// TIA Portal project "Project5" (V19)

(* hardware
DEVICE "S7-1500/ET200MP station_1"  S7-1500 station
   slot 0: "Rail_0"  Rack  6ES7 590-1***0-0AA0
   slot 1: "PLC_1"  CPU 1511C-1 PN  6ES7 511-1CK01-0AB0  V2.9
      slot 3: "CPU display_1"  6ES7591-1AA00-0AA0
      slot 32768: "PROFINET interface_1"  X1
         slot 32769: "Port_1"  X1 P1
         slot 32770: "Port_2"  X1 P2
      slot 34817: "Virtual CP interface port_1"  Virtual CP interface port  Virtual CP interface port
*)

// ===== PLC "PLC_1"  CPU 1511C-1 PN =====

VAR_GLOBAL   // PLC tag table "Default tag table"
   "Tag_1" AT %MW10 : Word;
   "Tag_2" AT %MD10 : DInt;
   "Tag_3" AT %MD20 : Real;
   "System_Byte" AT %MB100 : Byte;
   "FirstScan" AT %M100.0 : Bool;
   "DiagStatusUpdate" AT %M100.1 : Bool;
   "AlwaysTRUE" AT %M100.2 : Bool;
   "AlwaysFALSE" AT %M100.3 : Bool;
   "System_Byte(1)" AT %MB1 : Byte;
   "Clock_Byte" AT %MB100 : Byte;
   "Clock_10Hz" AT %M100.0 : Bool;
   "Clock_5Hz" AT %M100.1 : Bool;
   "Clock_2.5Hz" AT %M100.2 : Bool;
   "Clock_2Hz" AT %M100.3 : Bool;
   "Clock_1.25Hz" AT %M100.4 : Bool;
   "Clock_1Hz" AT %M100.5 : Bool;
   "Clock_0.625Hz" AT %M100.6 : Bool;
   "Clock_0.5Hz" AT %M100.7 : Bool;
   "Tag_4" AT %MW200 : Word;
   "Tag_5" AT %MW202 : Word;
   "Tag_6" AT %MD202 : Real;
END_VAR

DATA_BLOCK "FB_Motor_Speed_Calc_DB"   // DB1
{ S7_Optimized_Access := 'TRUE' }
VERSION : 0.1
// stored: InstanceOfName FB_Motor_Speed_Calc
"FB_Motor_Speed_Calc"
BEGIN
END_DATA_BLOCK

DATA_BLOCK "FB_Motor_Speed_Calc_Max_DB"   // DB3
{ S7_Optimized_Access := 'TRUE' }
VERSION : 0.2
// stored: InstanceOfName FB_Motor_Speed_Calc_Max
"FB_Motor_Speed_Calc_Max"
BEGIN
END_DATA_BLOCK

FUNCTION_BLOCK "FB_Motor_Speed_Calc"   // FB1, SCL
{ S7_Optimized_Access := 'TRUE' }
VERSION : 0.1
   VAR_INPUT
      Current_HSC_Count : DInt;   // Current value of the high-speed counter (e.g., LADDR#272)
      Run_Calculation : Bool;   // Trigger to run the calculation (e.g., driven by a 1s clock or OB35)
      Measurement_Interval_ms : Real := 1000.0;   // The fixed time interval for measurement (e.g., 1000.0 ms = 1 second)
      Pulses_Per_Revolution : Real := 1.0;   // Number of pulses generated by the sensor per one revolution (User specified 1)
   END_VAR
   VAR_OUTPUT
      RPM_Out : Real;   // Calculated motor speed in Revolutions Per Minute
   END_VAR
   VAR
      Previous_Count : DInt;   // Internal memory to store the count from the last calculation cycle (STATIC)
   END_VAR
   VAR_TEMP
      Time_Interval_s : Real;
      Delta_Count : Real;
   END_VAR
BEGIN
       // ----------------------------------------------------------------------
       // Speed Calculation Logic (Delta Count Method)
       // Runs only when the 'Run_Calculation' trigger is true (e.g., once every second)
       // Formula: RPM = (Delta_Count / Time_Interval_s) * (60.0 / PPR)
       // ----------------------------------------------------------------------

       IF #Run_Calculation THEN

           // 1. Calculate the change in count (Delta_Count)
           // DINT is used for counters. We convert to REAL for calculation accuracy.
           // We must handle the case where the counter may reset (Current < Previous),
           // although for modern PLCs reading a DINT HSC value, this is less likely 
           // to happen within a short interval.

           // Calculate the difference between the current count and the count from the last cycle

           // Check for potential counter rollover (Current_HSC_Count < Previous_Count)
           // If it rolls over, the difference will be negative, and the magnitude will be large,
           // but typically the HSC configuration handles this by resetting to 0. 
           // Assuming a standard incremental count:
           #Delta_Count := DINT_TO_REAL(#Current_HSC_Count -#Previous_Count);

           // 2. Convert the measurement interval from milliseconds to seconds
           #Time_Interval_s := #Measurement_Interval_ms / 1000.0;

           // 3. Check for division by zero (should not happen if Measurement_Interval_ms > 0)
           IF #Time_Interval_s > 0.0 AND #Pulses_Per_Revolution > 0.0 THEN

               // Calculate the speed in RPM
               // (Counts/second) * 60 = Counts/minute
               // (Counts/minute) / PPR = Revolutions/minute (RPM)
               #RPM_Out := (#Delta_Count / #Time_Interval_s) * (60.0 /#Pulses_Per_Revolution);

           ELSE
               #RPM_Out := 0.0;
           END_IF;

           // 4. Store the current count for the next calculation cycle
           #Previous_Count :=#Current_HSC_Count;

       END_IF;
END_FUNCTION_BLOCK

FUNCTION_BLOCK "FB_Motor_Speed_Calc_Max"   // FB2, SCL
{ S7_Optimized_Access := 'TRUE' }
VERSION : 0.2
   VAR_INPUT
      Current_HSC_Count : DInt;   // Current value of the high-speed counter
      Run_Calculation : Bool;   // Trigger to run the calculation (e.g., driven by a 1s clock or OB35)
      Reset_Max_RPM : Bool;   // New input: Use a momentary pulse to reset Max_RPM_Out to 0.0
      Measurement_Interval_ms : Real := 1000.0;   // The fixed time interval for measurement (e.g., 1000.0 ms = 1 second)
      Pulses_Per_Revolution : Real := 1.0;   // Number of pulses generated by the sensor per one revolution
   END_VAR
   VAR_OUTPUT
      RPM_Out : Real;   // Calculated current motor speed in Revolutions Per Minute
      Max_RPM_Out : Real;   // Output: Stores the highest RPM achieved since the last reset
   END_VAR
   VAR
      Previous_Count : DInt;   // Internal memory to store the count from the last calculation cycle (STATIC)
      s_Max_RPM_Value : Real;   // STATIC: Internal memory to persistently store the maximum RPM achieved. Initialized to 0.0 on creation.
   END_VAR
   VAR_TEMP
      Delta_Count : Real;
      Time_Interval_s : Real;
   END_VAR
BEGIN

       // ----------------------------------------------------------------------
       // 1. Reset Logic (Dominant)
       // If the Reset pulse is active, the internal maximum value is cleared.
       // ----------------------------------------------------------------------
       IF #Reset_Max_RPM THEN
           #s_Max_RPM_Value := 0.0;
       END_IF;

       // ----------------------------------------------------------------------
       // 2. Speed Calculation Logic (Runs only when the time trigger is true)
       // ----------------------------------------------------------------------
       IF #Run_Calculation THEN


           // Calculate the difference in counts over the interval
           #Delta_Count := DINT_TO_REAL(#Current_HSC_Count - #Previous_Count);

           // Convert the measurement interval from milliseconds to seconds
           #Time_Interval_s := #Measurement_Interval_ms / 1000.0;

           // Check for division by zero and calculate Current RPM
           IF #Time_Interval_s > 0.0 AND #Pulses_Per_Revolution > 0.0 THEN

               // Calculate Current RPM
               #RPM_Out := (#Delta_Count / #Time_Interval_s) * (60.0 /#Pulses_Per_Revolution);

               // 3. Maximum RPM Tracking Logic
               // If the currently calculated RPM is greater than the recorded internal maximum, update the internal maximum.
               IF #RPM_Out>#s_Max_RPM_Value THEN
                   #s_Max_RPM_Value:=#RPM_Out;
               END_IF;

           ELSE
               #RPM_Out := 0.0;
           END_IF;

           // Store the current count for the next calculation cycle
           #Previous_Count:=#Current_HSC_Count;

       END_IF;

       // ----------------------------------------------------------------------
       // 4. Output Assignment
       // Assign the internal persistent maximum value to the external output.
       // ----------------------------------------------------------------------
       #Max_RPM_Out := #s_Max_RPM_Value;
END_FUNCTION_BLOCK

ORGANIZATION_BLOCK "Main"   // OB1, LAD, ProgramCycle
TITLE = "Main Program Sweep (Cycle)"
{ S7_Optimized_Access := 'TRUE' }
VERSION : 0.1
   VAR_INPUT
      Initial_Call : Bool;   // Initial call of this OB
      Remanence : Bool;   // =True, if remanent data are available
   END_VAR
BEGIN

REGION Network 2
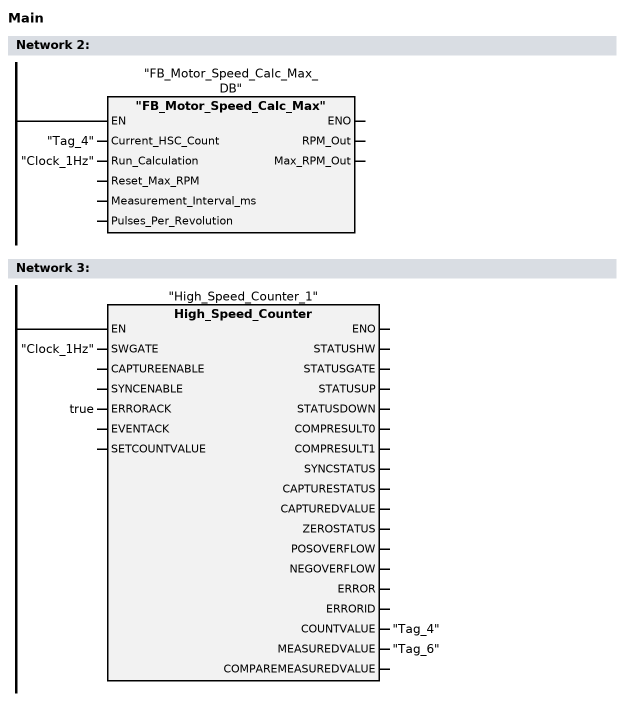
   RUNG wire#powerrail
      "FB_Motor_Speed_Calc_Max_DB"(Current_HSC_Count := "Tag_4", Run_Calculation := "Clock_1Hz", Reset_Max_RPM :=, Measurement_Interval_ms :=, Pulses_Per_Revolution :=, RPM_Out =>, Max_RPM_Out =>)
   END_RUNG
   // the same network as SCL:
   "FB_Motor_Speed_Calc_Max_DB"(Current_HSC_Count := "Tag_4", Run_Calculation := "Clock_1Hz");   // "FB_Motor_Speed_Calc_Max"
END_REGION

REGION Network 3
   "High_Speed_Counter_1"(SwGate := "Clock_1Hz",   // High_Speed_Counter
                          ErrorAck := true,
                          CountValue => "Tag_4",
                          MeasuredValue => "Tag_6");
END_REGION
END_ORGANIZATION_BLOCK